(* PLC project forms.project, CODESYS CODESYS V3.5 SP17 Patch 3 *)
(* stored: creationDateTime 2026-10-20T03:44:11.3191454, modificationDateTime 1601-01-01T03:00:00 *)

PROGRAM PRG_ProbeMain
  VAR
    fbOop : FB_ProbeOop;
  END_VAR

            fbOop(xIn := GVL_Probe.xFlag);
GVL_Probe.diHours := GVL_Probe.diHours + 1;

          
END_PROGRAM
